(* IEC 61131-3 sources: IRIS-Project/LASAL CONTROL SOFTWARE/LasalProject_2025_09_12/Network/IRIS_Manager, 1 file *)

(* ---- ONE_IRIS_MANAGER_Table.st ---- *)
#define OBJECTS_CONFIG

FUNCTION GLOBAL TAB ONE_IRIS_MANAGER
-1$UINT, 0$UINT,
0$UINT, 0$UINT,

11$UDINT,
TO_UDINT(2706637582), "Attuatore", 0$UINT, 0$UINT, 2$UINT,
TO_UDINT(1203230383), "MainSequence", 0$UINT, 0$UINT, 1$UINT,
TO_UDINT(3218456232), "Manager_globale", 0$UINT, 0$UINT, 1$UINT,
TO_UDINT(365955750), "ManagerMotori", 0$UINT, 0$UINT, 1$UINT,
TO_UDINT(2366454265), "Motore_M1", 0$UINT, 0$UINT, 1$UINT,
TO_UDINT(335833155), "Motore_M2", 0$UINT, 0$UINT, 1$UINT,
TO_UDINT(1661163733), "Motore_M3", 0$UINT, 0$UINT, 1$UINT,
TO_UDINT(4251438454), "Motore_M4", 0$UINT, 0$UINT, 1$UINT,
TO_UDINT(2321612256), "Motore_M5", 0$UINT, 0$UINT, 1$UINT,
TO_UDINT(325692506), "Motore_M6", 0$UINT, 0$UINT, 1$UINT,
TO_UDINT(1684970700), "Motore_M7", 0$UINT, 0$UINT, 1$UINT,

_NO_ATTR, TO_UDINT(1690670771), "ATTUATORE1",
_NO_ATTR, TO_UDINT(4258055945), "ATTUATORE2",

_NO_ATTR, TO_UDINT(3321030168), "MAINSEQUENCE1",

_NO_ATTR, TO_UDINT(1533940179), "MANAGER_GLOBALE1",

_NO_ATTR, TO_UDINT(3162257760), "MANAGERMOTORI1",

_NO_ATTR, TO_UDINT(1194371126), "MOTORE_M11",

_NO_ATTR, TO_UDINT(1813904373), "MOTORE_M21",

_NO_ATTR, TO_UDINT(1963379380), "MOTORE_M31",

_NO_ATTR, TO_UDINT(977755251), "MOTORE_M41",

_NO_ATTR, TO_UDINT(593259826), "MOTORE_M51",

_NO_ATTR, TO_UDINT(141639409), "MOTORE_M61",

_NO_ATTR, TO_UDINT(292163504), "MOTORE_M71",

//Internal connections
0$UDINT,
0$UDINT,
0$UDINT,
30$UDINT,
TO_UDINT(2), "Comando_manager_motori", TO_UDINT(4), "ClassSvr",
TO_UDINT(2), "Comando_manager_globale", TO_UDINT(3), "ClassSvr",
TO_UDINT(3), "Comando_main_sequence", TO_UDINT(2), "ClassSvr",
TO_UDINT(4), "M1_status", TO_UDINT(5), "ClassSvr",
TO_UDINT(4), "M1_command", TO_UDINT(5), "ClassSvr",
TO_UDINT(4), "M2_status", TO_UDINT(6), "ClassSvr",
TO_UDINT(4), "M2_command", TO_UDINT(6), "ClassSvr",
TO_UDINT(4), "M3_status", TO_UDINT(7), "ClassSvr",
TO_UDINT(4), "M3_command", TO_UDINT(7), "ClassSvr",
TO_UDINT(4), "M4_status", TO_UDINT(8), "ClassSvr",
TO_UDINT(4), "M4_command", TO_UDINT(8), "ClassSvr",
TO_UDINT(4), "M5_status", TO_UDINT(9), "ClassSvr",
TO_UDINT(4), "M5_command", TO_UDINT(9), "ClassSvr",
TO_UDINT(4), "M6_status", TO_UDINT(10), "ClassSvr",
TO_UDINT(4), "M6_command", TO_UDINT(10), "ClassSvr",
TO_UDINT(4), "Homing_complete", TO_UDINT(2), "ClassSvr",
TO_UDINT(4), "Phasing_complete", TO_UDINT(2), "ClassSvr",
TO_UDINT(4), "Charge_complete", TO_UDINT(2), "ClassSvr",
TO_UDINT(4), "Irradiation_complete", TO_UDINT(2), "ClassSvr",
TO_UDINT(4), "Discharge_complete", TO_UDINT(2), "ClassSvr",
TO_UDINT(4), "Stop_client", TO_UDINT(2), "ClassSvr",
TO_UDINT(4), "ToManagerGlobale", TO_UDINT(3), "ClassSvr",
TO_UDINT(4), "c_1_3_pelletMode_M2", TO_UDINT(6), "s_1_3_pelletMode",
TO_UDINT(4), "c_1_3_pelletMode_M4", TO_UDINT(8), "s_1_3_pelletMode",
TO_UDINT(4), "c_1_3_pelletMode_M5", TO_UDINT(9), "s_1_3_pelletMode",
TO_UDINT(4), "c_PelletAvailable", TO_UDINT(9), "ClassSvr",
TO_UDINT(8), "Comando_to_M8Class", TO_UDINT(11), "ClassSvr",
TO_UDINT(9), "Comando_Attuatore_1", TO_UDINT(0), "ClassSvr",
TO_UDINT(9), "Comando_Attuatore_2", TO_UDINT(1), "ClassSvr",
TO_UDINT(11), "Stato_to_M4", TO_UDINT(8), "ClassSvr",

//Initialization values
0$UDINT,
7$UDINT,
TO_UDINT(0), "R_p", TO_UDINT(0),//|IRIS_MANAGER.Attuatore1.R_p;
TO_UDINT(0), "R_aus_1", TO_UDINT(0),//|IRIS_MANAGER.Attuatore1.R_aus_1;
TO_UDINT(0), "R_aus_2", TO_UDINT(0),//|IRIS_MANAGER.Attuatore1.R_aus_2;
TO_UDINT(1), "R_p", TO_UDINT(0),//|IRIS_MANAGER.Attuatore2.R_p;
TO_UDINT(1), "R_aus_1", TO_UDINT(0),//|IRIS_MANAGER.Attuatore2.R_aus_1;
TO_UDINT(1), "R_aus_2", TO_UDINT(0),//|IRIS_MANAGER.Attuatore2.R_aus_2;
TO_UDINT(5), "Comando_M1", TO_UDINT(PASSIVE_LMCAXIS),//|IRIS_MANAGER.Motore_M11.Comando_M1;

//Symbolic initialization values
0$UDINT,
0$UDINT,

//Initialization of string values
0$UDINT,
0$UDINT,

//Configuration of tasks (RealTime, Cyclic, Background)
0$UDINT,
0$UDINT,

0$UDINT,
12$UDINT,
TO_UDINT(0), (100)$UDINT, 4194303$DINT, 	//ATTUATORE1
TO_UDINT(1), (100)$UDINT, 4194303$DINT, 	//ATTUATORE2
TO_UDINT(2), (100)$UDINT, 4194303$DINT, 	//MAINSEQUENCE1
TO_UDINT(3), (100)$UDINT, 4194303$DINT, 	//MANAGER_GLOBALE1
TO_UDINT(4), (100)$UDINT, 4194303$DINT, 	//MANAGERMOTORI1
TO_UDINT(5), (100)$UDINT, 4194303$DINT, 	//MOTORE_M11
TO_UDINT(6), (100)$UDINT, 4194303$DINT, 	//MOTORE_M21
TO_UDINT(7), (100)$UDINT, 4194303$DINT, 	//MOTORE_M31
TO_UDINT(8), (100)$UDINT, 4194303$DINT, 	//MOTORE_M41
TO_UDINT(9), (100)$UDINT, 4194303$DINT, 	//MOTORE_M51
TO_UDINT(10), (100)$UDINT, 4194303$DINT, 	//MOTORE_M61
TO_UDINT(11), (100)$UDINT, 4194303$DINT, 	//MOTORE_M71

0$UDINT,
0$UDINT,

//External connections
0$UDINT,
47$UDINT,
TO_UDINT(0), "R_p", C_DIR, TO_UDINT(1390357230), "TO1271","Output1",
TO_UDINT(0), "R_aus_1", C_DIR, TO_UDINT(1390357230), "TO1271","Output2",
TO_UDINT(0), "R_aus_2", C_DIR, TO_UDINT(1390357230), "TO1271","Output3",
TO_UDINT(1), "R_p", C_DIR, TO_UDINT(1390357230), "TO1271","Output5",
TO_UDINT(1), "R_aus_1", C_DIR, TO_UDINT(1390357230), "TO1271","Output6",
TO_UDINT(1), "R_aus_2", C_DIR, TO_UDINT(1390357230), "TO1271","Output7",
TO_UDINT(3), "Reset_IN", C_TRY, TO_UDINT(2516706254), "DI1601","Input3",
TO_UDINT(3), "c_ResetTimer", C_DIR, TO_UDINT(1081583723), "Reset1","s_ResetT",
TO_UDINT(4), "LED_Rosso", C_DIR, TO_UDINT(1390357230), "TO1271","Output8",
TO_UDINT(4), "LED_Arancione", C_DIR, TO_UDINT(1390357230), "TO1271","Output11",
TO_UDINT(4), "LED_Verde", C_DIR, TO_UDINT(1390357230), "TO1271","Output10",
TO_UDINT(4), "c_MPS_Req", C_DIR, TO_UDINT(3838738401), "MPS1","ReqToMPS",
TO_UDINT(4), "c_1_3_pelletMode_TimerMov", C_DIR, TO_UDINT(136251601), "MoveTimer1","s_1_3_pelletMode",
TO_UDINT(4), "c_1_3_pelletMode_TimerIrr", C_DIR, TO_UDINT(101499717), "IrradiationTimers","s_1_3_pelletMode",
TO_UDINT(5), "Comando_M1", C_TRY, TO_UDINT(1906010274), "_LMCAxis_M1","Control",
TO_UDINT(5), "M1_LS_1", C_DIR, TO_UDINT(201264582), "ST1511","Input1",
TO_UDINT(5), "M1_LS_2", C_TRY, TO_UDINT(201264582), "ST1511","Input2",
TO_UDINT(5), "c_MaxCurrent", C_DIR, TO_UDINT(201264582), "ST1511","MaxCurrent",
TO_UDINT(5), "SetPosition_Controller", C_DIR, TO_UDINT(1906010274), "_LMCAxis_M1","ActPos",
TO_UDINT(6), "Comando_M2", C_DIR, TO_UDINT(3901896984), "_LMCAxis_M2","Control",
TO_UDINT(6), "M2_LS", C_TRY, TO_UDINT(2465619068), "ST1512","Input2",
TO_UDINT(6), "SetPosition_Controller", C_DIR, TO_UDINT(3901896984), "_LMCAxis_M2","ActPos",
TO_UDINT(7), "Comando_M3", C_DIR, TO_UDINT(2677344654), "_LMCAxis_M3","Control",
TO_UDINT(7), "M3_LS_1", C_TRY, TO_UDINT(3857804522), "ST1513","Input1",
TO_UDINT(7), "M3_LS_2", C_TRY, TO_UDINT(3857804522), "ST1513","Input2",
TO_UDINT(7), "c_MaxCurrent", C_DIR, TO_UDINT(3857804522), "ST1513","MaxCurrent",
TO_UDINT(7), "SetPositionController", C_DIR, TO_UDINT(2677344654), "_LMCAxis_M3","ActPos",
TO_UDINT(8), "Comando_M4", C_DIR, TO_UDINT(32611373), "_LMCAxis_M4","Control",
TO_UDINT(8), "M4_LS", C_TRY, TO_UDINT(2073426249), "ST1514","Input1",
TO_UDINT(8), "c_MaxCurrent", C_DIR, TO_UDINT(2073426249), "ST1514","MaxCurrent",
TO_UDINT(8), "SetPositionController", C_DIR, TO_UDINT(32611373), "_LMCAxis_M4","ActPos",
TO_UDINT(8), "c_TimerDis", C_TRY, TO_UDINT(4223322087), "DischargeTimer1","s_StartStopTimer",
TO_UDINT(8), "c_TimerMov", C_DIR, TO_UDINT(136251601), "MoveTimer1","s_StartStopTimer",
TO_UDINT(9), "Comando_M5", C_DIR, TO_UDINT(1995877563), "_LMCAxis_M5","Control",
TO_UDINT(9), "M5_LS", C_TRY, TO_UDINT(210946527), "ST1515","Input1",
TO_UDINT(9), "c_MaxCurrent", C_DIR, TO_UDINT(210946527), "ST1515","MaxCurrent",
TO_UDINT(9), "SetPosition_Controller", C_DIR, TO_UDINT(1995877563), "_LMCAxis_M5","ActPos",
TO_UDINT(9), "c_TimerMov", C_DIR, TO_UDINT(136251601), "MoveTimer1","s_StartStopTimer",
TO_UDINT(9), "c_TimerIrr", C_DIR, TO_UDINT(101499717), "IrradiationTimers","s_TimerStartStop",
TO_UDINT(10), "Comando_M6", C_DIR, TO_UDINT(4026531073), "_LMCAxis_M6","Control",
TO_UDINT(10), "M6_LS_1", C_TRY, TO_UDINT(2510002277), "ST1516","Input1",
TO_UDINT(10), "M6_LS_2", C_TRY, TO_UDINT(2510002277), "ST1516","Input2",
TO_UDINT(10), "SetPosition_Controller", C_DIR, TO_UDINT(4026531073), "_LMCAxis_M6","ActPos",
TO_UDINT(11), "Comando_M7", C_DIR, TO_UDINT(2566442391), "_LMCAxis_M7","Control",
TO_UDINT(11), "M7_LS_1", C_TRY, TO_UDINT(3801917683), "ST1517","Input1",
TO_UDINT(11), "M7_LS_2", C_TRY, TO_UDINT(3801917683), "ST1517","Input2",
TO_UDINT(11), "SetPositionController", C_DIR, TO_UDINT(2566442391), "_LMCAxis_M7","ActPos",

//Magic internal connections
0$UDINT,
0$UDINT,

//Configuration of timeslots of tasks (RealTime, Cyclic)
#ifdef __LSLLDR_TIMESLOTS__
0$UDINT,
0$UDINT,

0$UDINT,
0$UDINT,

#endif //__LSLLDR_TIMESLOTS__

//MultiMaster connections
#ifdef __LSLLDR_MULTIMASTER__
0$UDINT,
0$UDINT,
#endif //__LSLLDR_MULTIMASTER__

//Configuration for task ID (RealTime, CyclicTime)
#ifdef __LSLLDR_TASKID__
"\\\\TASKS2  "
0$UDINT,
0$UDINT,

0$UDINT,
12$UDINT,
(0)$UDINT, 	//ATTUATORE1
(0)$UDINT, 	//ATTUATORE2
(0)$UDINT, 	//MAINSEQUENCE1
(0)$UDINT, 	//MANAGER_GLOBALE1
(0)$UDINT, 	//MANAGERMOTORI1
(0)$UDINT, 	//MOTORE_M11
(0)$UDINT, 	//MOTORE_M21
(0)$UDINT, 	//MOTORE_M31
(0)$UDINT, 	//MOTORE_M41
(0)$UDINT, 	//MOTORE_M51
(0)$UDINT, 	//MOTORE_M61
(0)$UDINT, 	//MOTORE_M71

0$UDINT,
0$UDINT,

#endif //__LSLLDR_TASKID__

END_FUNCTION
